SUBAPPLICATION Ventilsteuerung (* Subapplication Type *)
  (* Standard: 61499-2 *)
  (* Version 1.0, 2023-10-23, franz *)
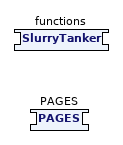
  SUBAPPS
    functions : SlurryTanker;
    PAGES : PAGES;
  END_SUBAPPS
END_SUBAPPLICATION
